(* IEC 61131-3 sources: rusty/tests/lit/single/type_promotion/constants, 3 files *)

(* ---- initializer_from_other_signedness.st ---- *)
// RUN: %COMPILE %s && %RUN | %CHECK %s
// XFAIL: *
// A constant initialized from a constant of other signedness is extended by the signedness of the target, not of the source.
VAR_GLOBAL CONSTANT
    cu : USINT := 200;
    k : INT := cu;
    cs : SINT := -1;
    u : ULINT := cs;
    d : DINT := cs;
END_VAR

VAR_GLOBAL
    g : INT := cu;
END_VAR

FUNCTION main : DINT
    VAR CONSTANT
        lk : INT := cu;
    END_VAR
    VAR
        t : INT := USINT#200;
    END_VAR

    printf('variable INT := USINT 200 = %d$N', g);          // CHECK: variable INT := USINT 200 = 200
    printf('constant INT := USINT 200 = %d$N', k);          // CHECK-NEXT: constant INT := USINT 200 = 200
    printf('local constant INT := USINT 200 = %d$N', lk);   // CHECK-NEXT: local constant INT := USINT 200 = 200
    printf('INT := USINT#200 = %d$N', t);                   // CHECK-NEXT: INT := USINT#200 = 200
    printf('constant ULINT := SINT -1 = %llu$N', u);        // CHECK-NEXT: constant ULINT := SINT -1 = 18446744073709551615
    printf('constant DINT := SINT -1 = %d$N', d);           // CHECK-NEXT: constant DINT := SINT -1 = -1
END_FUNCTION

(* ---- overflowing_initializer.st ---- *)
// RUN: %COMPILE %s && %RUN | %CHECK %s
// XFAIL: *
// A global constant whose initializer overflows its type aborts code generation.
VAR_GLOBAL CONSTANT
    c1 : USINT := 200;
    c2 : SINT := 0 - c1;
END_VAR

VAR_GLOBAL
    g : SINT := 0 - c1;
END_VAR

FUNCTION main : DINT
    printf('variable SINT := 0 - 200 = %d$N', g);           // CHECK: variable SINT := 0 - 200 = 56
    printf('constant SINT := 0 - 200 = %d$N', c2);          // CHECK-NEXT: constant SINT := 0 - 200 = 56
END_FUNCTION

(* ---- unsigned_constant_operands.st ---- *)
// RUN: %COMPILE %s && %RUN | %CHECK %s
// Compares, divisions and MOD on UDINT constants follow the same unsigned rules as on variables.
VAR_GLOBAL CONSTANT
    big : UDINT := 4000000000;
    small : UDINT := 5;
END_VAR

VAR_GLOBAL
    half : UDINT := big / 2;
    rest : UDINT := big MOD 7;
END_VAR

FUNCTION main : DINT
    VAR
        q : UDINT;
    END_VAR

    // Folded initializers
    printf('initializer big / 2 = %u$N', half);             // CHECK: initializer big / 2 = 2000000000
    printf('initializer big MOD 7 = %u$N', rest);           // CHECK-NEXT: initializer big MOD 7 = 3

    // Body expressions on constants
    q := big / 2;
    printf('body big / 2 = %u$N', q);                       // CHECK-NEXT: body big / 2 = 2000000000
    printf('big > small = %d$N', big > small);              // CHECK-NEXT: big > small = 1
    printf('big > 5 = %d$N', big > 5);                      // CHECK-NEXT: big > 5 = 1
END_FUNCTION
